// TIA Portal project "Coffee maker machine" (V14)

(* hardware
DEVICE "S7-1200 station_1"  S7-1200 Station
   slot 0: "Rack_0"  S7-1200 Rack  Rack  V1.0
   slot 1: "PLC_1"  CPU 1215C DC/DC/Rly  6ES7 215-1HG40-0XB0  V4.0
*)

// ===== PLC "PLC_1"  CPU 1215C DC/DC/Rly =====

VAR_GLOBAL   // PLC tag table "Default tag table"
   "START" AT %I0.0 : Bool;
   "STOP" AT %I0.1 : Bool;
   "PROCESS" AT %M0.0 : Bool;
   "coin" AT %I0.2 : Bool;
   "CUP" AT %Q0.0 : Bool;
   "COFFEE VALVE" AT %Q0.1 : Bool;
   "HW VALVE" AT %Q0.2 : Bool;
   "MIXING CHMBR" AT %Q0.3 : Bool;
   "TUANG KOPI" AT %Q0.4 : Bool;
   "KOPI HABIS" AT %Q0.5 : Bool;
   "BUBUK HABIS" AT %Q0.6 : Bool;
   "AIR HABIS" AT %Q0.7 : Bool;
   "RST CUP" AT %I0.3 : Bool;
   "RST BUBUK" AT %I0.4 : Bool;
   "RST AIR" AT %I0.5 : Bool;
END_VAR

// folder: System blocks/Program resources

DATA_BLOCK "PC OUTLET"   // DB1
{ S7_Optimized_Access := 'TRUE' }
AUTHOR : Simatic
FAMILY : IEC
NAME : IEC_TMR
VERSION : 1.0
// stored: InstanceOfName IEC_TIMER
"IEC_TIMER"
BEGIN
END_DATA_BLOCK

DATA_BLOCK "COFFEE_HW"   // DB2
{ S7_Optimized_Access := 'TRUE' }
AUTHOR : Simatic
FAMILY : IEC
NAME : IEC_TMR
VERSION : 1.0
// stored: InstanceOfName IEC_TIMER
"IEC_TIMER"
BEGIN
END_DATA_BLOCK

DATA_BLOCK "MIXING"   // DB3
{ S7_Optimized_Access := 'TRUE' }
AUTHOR : Simatic
FAMILY : IEC
NAME : IEC_TMR
VERSION : 1.0
// stored: InstanceOfName IEC_TIMER
"IEC_TIMER"
BEGIN
END_DATA_BLOCK

DATA_BLOCK "POUR VALVE"   // DB4
{ S7_Optimized_Access := 'TRUE' }
AUTHOR : Simatic
FAMILY : IEC
NAME : IEC_TMR
VERSION : 1.0
// stored: InstanceOfName IEC_TIMER
"IEC_TIMER"
BEGIN
END_DATA_BLOCK

DATA_BLOCK "counter"   // DB5
{ S7_Optimized_Access := 'TRUE' }
AUTHOR : Simatic
FAMILY : IEC
NAME : CNTR
VERSION : 1.0
// stored: InstanceOfName IEC_COUNTER
"IEC_COUNTER"
BEGIN
END_DATA_BLOCK

DATA_BLOCK "CounterBUBUK"   // DB6
{ S7_Optimized_Access := 'TRUE' }
AUTHOR : Simatic
FAMILY : IEC
NAME : CNTR
VERSION : 1.0
// stored: InstanceOfName IEC_COUNTER
"IEC_COUNTER"
BEGIN
END_DATA_BLOCK

DATA_BLOCK "counterAIR"   // DB7
{ S7_Optimized_Access := 'TRUE' }
AUTHOR : Simatic
FAMILY : IEC
NAME : CNTR
VERSION : 1.0
// stored: InstanceOfName IEC_COUNTER
"IEC_COUNTER"
BEGIN
END_DATA_BLOCK

// folder: (top level)

ORGANIZATION_BLOCK "Main"   // OB1, LAD, ProgramCycle
TITLE = "Main Program Sweep (Cycle)"
{ S7_Optimized_Access := 'TRUE' }
VERSION : 0.1
   VAR_INPUT
      Initial_Call : Bool;   // Initial call of this OB
      Remanence : Bool;   // =True, if remanent data are available
   END_VAR
BEGIN

REGION Network 1
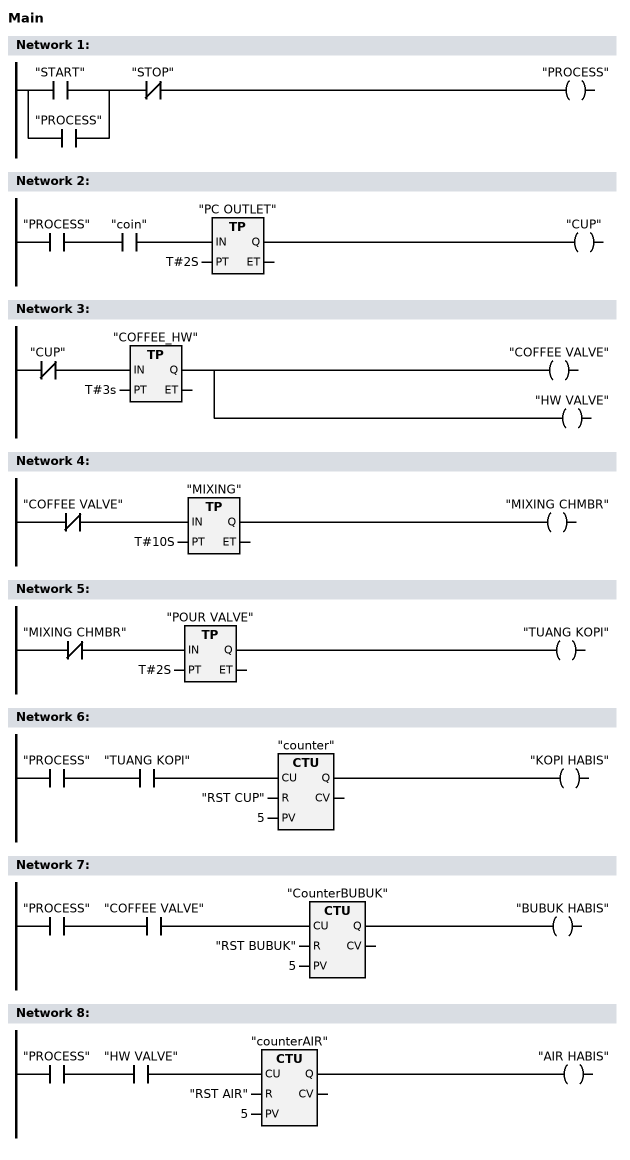
   RUNG wire#powerrail
      Contact( "START" )
      wire#w1
      I_Contact( "STOP" )
      Coil( "PROCESS" )
   END_RUNG
   RUNG wire#powerrail
      Contact( "PROCESS" )
   END_RUNG wire#w1
   // the same network as SCL:
   "PROCESS" := ("START" OR "PROCESS") AND NOT "STOP";
END_REGION

REGION Network 2
   "PC OUTLET".TP(IN := "PROCESS" AND "coin", PT := T#2S);
   "CUP" := "PC OUTLET".Q;
END_REGION

REGION Network 3
   "COFFEE_HW".TP(IN := NOT "CUP", PT := T#3s);
   "COFFEE VALVE" := "COFFEE_HW".Q;
   "HW VALVE" := "COFFEE_HW".Q;
END_REGION

REGION Network 4
   "MIXING".TP(IN := NOT "COFFEE VALVE", PT := T#10S);
   "MIXING CHMBR" := "MIXING".Q;
END_REGION

REGION Network 5
   "POUR VALVE".TP(IN := NOT "MIXING CHMBR", PT := T#2S);
   "TUANG KOPI" := "POUR VALVE".Q;
END_REGION

REGION Network 6
   "counter".CTU(CU := "PROCESS" AND "TUANG KOPI", R := "RST CUP", PV := 5);
   "KOPI HABIS" := "counter".Q;
END_REGION

REGION Network 7
   "CounterBUBUK".CTU(CU := "PROCESS" AND "COFFEE VALVE", R := "RST BUBUK", PV := 5);
   "BUBUK HABIS" := "CounterBUBUK".Q;
END_REGION

REGION Network 8
   "counterAIR".CTU(CU := "PROCESS" AND "HW VALVE", R := "RST AIR", PV := 5);
   "AIR HABIS" := "counterAIR".Q;
END_REGION
END_ORGANIZATION_BLOCK